// TIA Portal project "PLC_4_LINE4" (V18)

(* hardware
DEVICE "S7-1500/ET200MP station_1"  S7-1500 station
   slot 0: "Rail_0"  Rack  6ES7 590-1***0-0AA0
   slot 1: "PLC_4"  CPU 1511-1 PN  6ES7 511-1AK02-0AB0  V2.9
      slot 3: "CPU display_1"  6ES7591-1AA00-0AA0
      slot 32768: "PROFINET interface_1"  X1
         slot 32769: "Port_1"  X1 P1
         slot 32770: "Port_2"  X1 P2
      slot 34817: "Virtual CP interface port_1"  Virtual CP interface port  Virtual CP interface port
   slot 2: "DI 32x24VDC HF_1"  DI 32x24VDC HF  6ES7 521-1BL00-0AB0  V2.2
   slot 3: "DI 32x24VDC HF_2"  DI 32x24VDC HF  6ES7 521-1BL00-0AB0  V2.2
   slot 4: "DQ 32x24VDC/0.5A HF_1"  DQ 32x24VDC/0.5A HF  6ES7 522-1BL01-0AB0  V1.1
*)

// ===== PLC "PLC_4"  CPU 1511-1 PN =====

VAR_GLOBAL   // PLC tag table "Default tag table"
   "Tag_1" AT %I0.3 : Bool;
   "Tag_2" AT %I0.4 : Bool;
   "Tag_3" AT %I0.5 : Bool;
   "Tag_4" AT %I0.0 : Bool;
   "Tag_5" AT %I0.1 : Bool;
   "Tag_6" AT %I2.1 : Bool;
   "Tag_7" AT %I0.7 : Bool;
   "Tag_8" AT %I1.6 : Bool;
   "Tag_9" AT %I1.0 : Bool;
   "Tag_10" AT %I1.1 : Bool;
   "Tag_11" AT %I1.2 : Bool;
   "Tag_12" AT %I1.3 : Bool;
   "Tag_13" AT %I1.4 : Bool;
   "Tag_14" AT %I1.5 : Bool;
   "Tag_15" AT %Q0.4 : Bool;
   "Tag_16" AT %Q0.5 : Bool;
   "Tag_17" AT %Q0.6 : Bool;
   "Tag_18" AT %Q0.7 : Bool;
   "Tag_19" AT %I4.3 : Bool;
   "Tag_20" AT %I4.4 : Bool;
   "Tag_21" AT %I4.5 : Bool;
   "Tag_22" AT %I4.0 : Bool;
   "Tag_23" AT %I4.1 : Bool;
   "Tag_24" AT %I6.1 : Bool;
   "Tag_25" AT %I4.7 : Bool;
   "Tag_26" AT %I4.6 : Bool;
   "Tag_27" AT %I5.0 : Bool;
   "Tag_28" AT %I5.1 : Bool;
   "Tag_29" AT %I5.2 : Bool;
   "Tag_30" AT %I5.3 : Bool;
   "Tag_31" AT %I5.4 : Bool;
   "Tag_32" AT %I5.5 : Bool;
   "Tag_33" AT %Q2.4 : Bool;
   "Tag_34" AT %Q2.5 : Bool;
   "Tag_35" AT %Q2.6 : Bool;
   "Tag_36" AT %Q2.7 : Bool;
END_VAR

TYPE "typeTask"
   STRUCT
      station : Int;
      dwell_s : Int;
      crane : String[4];
      tank_name : String[10];
      prev : Int;
      next : Int;
      status : Int;
   END_STRUCT;
END_TYPE

TYPE "typeCraneData"
   STRUCT
      task_count : Int;
      tasks : Array[1..20] of "typeTask";
      cmd_send : Bool;
      sts_busy : Bool;
      sts_done : Bool;
      sts_step : Int;
      sts_state : Int;
      ls_at : Array[0..20] of Bool;
      ls_dip : Bool;
      ls_up : Bool;
      ls_mid : Bool;
      btn_start : Bool;
      mv_fwd : Bool;
      mv_rev : Bool;
      mv_up : Bool;
      mv_down : Bool;
      estop : Bool;
      auto : Bool;
      cmd_reset : Bool;
      cmd_stop : Bool;
      pos : Array[0..20] of Int;
   END_STRUCT;
END_TYPE

DATA_BLOCK "Crane6Data"   // DB1
{ S7_Optimized_Access := 'TRUE' }
VERSION : 0.1
BEGIN
   pos[0] := 21;
   pos[1] := 20;
   pos[12] := 14;
   pos[13] := 15;
   pos[14] := 16;
   pos[15] := 17;
   pos[16] := 18;
   pos[17] := 19;
   pos[18] := 20;
END_DATA_BLOCK

DATA_BLOCK "Crane7AData"   // DB2
{ S7_Optimized_Access := 'TRUE' }
VERSION : 0.1
BEGIN
   pos[0] := 2;
   pos[1] := 1;
   pos[2] := 3;
   pos[3] := 4;
   pos[4] := 5;
   pos[5] := 6;
   pos[6] := 7;
   pos[7] := 8;
END_DATA_BLOCK

DATA_BLOCK "Crane6_Seq_DB"   // DB3
{ S7_Optimized_Access := 'TRUE' }
VERSION : 0.1
// stored: InstanceOfName CraneSequencer
"CraneSequencer"
BEGIN
END_DATA_BLOCK

DATA_BLOCK "Crane7A_Seq_DB"   // DB4
{ S7_Optimized_Access := 'TRUE' }
VERSION : 0.1
// stored: InstanceOfName CraneSequencer
"CraneSequencer"
BEGIN
END_DATA_BLOCK

FUNCTION_BLOCK "CraneSequencer"   // FB1, SCL
{ S7_Optimized_Access := 'TRUE' }
VERSION : 0.1
   VAR_IN_OUT
      d : "typeCraneData";
   END_VAR
   VAR
      state : Int;
      idx : Int;
      count : Int;
      cur : Int;
      prevSend : Bool;
      tHold : TON_TIME;
      tDwell : TON_TIME;
   END_VAR
   VAR_TEMP
      target : Int;
      arrived : Bool;
   END_VAR
BEGIN
   // ============================================================================
   //  CraneSequencer  —  GENERIC per-crane batch sequencer  (LIBRARY block)
   // ----------------------------------------------------------------------------
   //  ONE function block reused by EVERY crane on EVERY PLC. Call once per scan
   //  from OB1, passing that crane's data block as the InOut #d. No copy, no
   //  find/replace — the crane it drives is chosen entirely by which DB you pass.
   //
   //  Block type : FUNCTION BLOCK (FB), language SCL.
   //  InOut      : d : "typeCraneData"           // the whole crane interface (a DB of this UDT)
   //  Static     : state:Int, idx:Int, count:Int, cur:Int, prevSend:Bool,
   //               tHold:TON_TIME, tDwell:TON_TIME
   //  Temp       : target:Int, arrived:Bool
   //
   //  OB1 (per crane):  CraneSequencer(d := "Crane6Data")   // its own instance DB
   //                    CraneSequencer(d := "Crane7AData")
   //
   //  Stations: 0=Parking  1=Loading  2..N = tanks (tank number + 1).
   //  States : 0 IDLE · 10 GO_LOAD · 20 LOWER_LOAD · 30 WAIT_BTN · 40 LIFT_LOAD
   //           50 GO_TANK · 60 LOWER_TANK · 70 DWELL · 80 LIFT_TANK · 85 GO_PARK · 90 DONE
   //
   //  DIRECTION IS BY PHYSICAL POSITION, NOT STATION NUMBER.
   //  The plant is NOT laid out in station-number order: Parking sits WEST of Loading, and a
   //  downstream crane's Loading is a transfer tank at the far (West) end. So travel direction
   //  is decided from #d.pos[station] — the physical left→right position of each station
   //  (1 = East-most … larger = further West). TravelTo drives WEST (mv_fwd → R-West) toward a
   //  HIGHER pos, EAST (mv_rev → R-East) toward a LOWER pos. The station's arrival switch is still
   //  #d.ls_at[station]. **Set #d.pos[] per crane** — see the PLC's position-map doc.
   //
   //  COMMANDS (app/Manager writes these):
   //    cmd_send  — arm a batch (rising edge, from IDLE).
   //    cmd_stop  — EMERGENCY HOLD: kills all motion immediately, latches state 100 (STOPPED).
   //                Does NOT clear the recipe. Clear it (and Reset) to move again.
   //    cmd_reset — CLEAN/HOME: lift clear → travel to Parking → wipe the recipe → IDLE.
   //                "As if no recipe was sent, crane back at its home." PLC clears cmd_reset when done.
   //  Extra states: 100 STOPPED · 110 RESET_LIFT · 120 RESET_HOME.
   // ============================================================================

   // ---- command overrides (run BEFORE the state machine, highest priority) ----
   IF #d.cmd_stop THEN                       // immediate emergency hold (latched)
       #d.mv_fwd := FALSE;
       #d.mv_rev := FALSE;
       #d.mv_up := FALSE;
       #d.mv_down := FALSE;
       #d.sts_busy := FALSE;
       #state := 100;
   ELSIF #d.cmd_reset AND #state <> 110 AND #state <> 120 THEN   // start homing/clear (if not already)
       // Wipe the recipe IMMEDIATELY (visible at once), then home the crane.
       #d.task_count := 0;
       #d.sts_step := 0;
       #d.sts_done := FALSE;
       #d.cmd_send := FALSE;
       #idx := 0;
       #count := 0;
       #d.sts_busy := TRUE;
       #state := 110;
   END_IF;

   #d.sts_state := #state;

   CASE #state OF
       0:  // IDLE — parked, hoist up, motors off, waiting for a batch.
           #d.mv_fwd := FALSE;
           #d.mv_rev := FALSE;
           #d.mv_up := FALSE;
           #d.mv_down := FALSE;
           #d.sts_busy := FALSE;
           #d.sts_step := 0;
           IF #d.cmd_send AND NOT #prevSend AND #d.task_count > 0 THEN
               #count := #d.task_count;
               #idx := 1;
               #d.sts_done := FALSE;
               #d.sts_busy := TRUE;
               #state := 10;
           END_IF;

       10: // GO_LOAD — travel to the Loading Area (station 1).
           #d.sts_busy := TRUE;
           #target := 1;
           #arrived := "TravelTo"(target := #d.pos[#target], cur := #d.pos[#cur],
                                  atTarget := #d.ls_at[#target],
                                  fwd => #d.mv_fwd, rev => #d.mv_rev);
           IF #arrived THEN
               #cur := #target;
               #d.mv_fwd := FALSE;
               #d.mv_rev := FALSE;
               #state := 20;
           END_IF;

       20: // LOWER_LOAD — lower the hoist until the dip limit switch is made.
           #d.mv_up := FALSE;
           #d.mv_down := TRUE;
           IF #d.ls_dip THEN
               #d.mv_down := FALSE;
               #state := 30;
           END_IF;

       30: // WAIT_BTN — operator loads material, then HOLDS btn_start for 3 s.
           #tHold(IN := #d.btn_start,
                  PT := T#3S);
           IF #tHold.Q THEN
               #state := 40;
           END_IF;

       40: // LIFT_LOAD — raise the hoist clear before travelling.
           #d.mv_down := FALSE;
           #d.mv_up := TRUE;
           IF #d.ls_up THEN
               #d.mv_up := FALSE;
               #state := 50;
           END_IF;

       50: // GO_TANK — travel to THIS task's tank station (TravelTo reverses if lower).
           #d.sts_step := #idx;
           #d.tasks[#idx].status := 1;                  // running
           #target := #d.tasks[#idx].station;
           #arrived := "TravelTo"(target := #d.pos[#target], cur := #d.pos[#cur],
                                  atTarget := #d.ls_at[#target],
                                  fwd => #d.mv_fwd, rev => #d.mv_rev);
           IF #arrived THEN
               #cur := #target;
               #d.mv_fwd := FALSE;
               #d.mv_rev := FALSE;
               #state := 60;
           END_IF;

       60: // LOWER_TANK — dip into the tank until the dip limit switch is made.
           #d.mv_up := FALSE;
           #d.mv_down := TRUE;
           IF #d.ls_dip THEN
               #d.mv_down := FALSE;
               #state := 70;
           END_IF;

       70: // DWELL — hold in the tank for this task's dwell_s seconds.
           #tDwell(IN := TRUE,
                   PT := DINT_TO_TIME(INT_TO_DINT(#d.tasks[#idx].dwell_s) * 1000));
           IF #tDwell.Q THEN
               #tDwell(IN := FALSE,
                       PT := T#0S);        // reset the timer for the next tank
               #state := 80;
           END_IF;

       80: // LIFT_TANK — lift out, mark the task done, advance or finish.
           #d.mv_down := FALSE;
           #d.mv_up := TRUE;
           IF #d.ls_up THEN
               #d.mv_up := FALSE;
               #d.tasks[#idx].status := 2;              // done
               IF #idx < #count THEN
                   #idx := #idx + 1;
                   #state := 50;                        // next tank
               ELSE
                   #state := 85;                        // all tanks done
               END_IF;
           END_IF;

       85: // GO_PARK — return home to Parking (station 0).
           #target := 0;
           #arrived := "TravelTo"(target := #d.pos[#target], cur := #d.pos[#cur],
                                  atTarget := #d.ls_at[#target],
                                  fwd => #d.mv_fwd, rev => #d.mv_rev);
           IF #arrived THEN
               #cur := #target;
               #d.mv_fwd := FALSE;
               #d.mv_rev := FALSE;
               #state := 90;
           END_IF;

       90: // DONE — raise the done flag, wait for the app to acknowledge (cmd_send → FALSE).
           #d.sts_busy := FALSE;
           #d.sts_done := TRUE;
           IF NOT #d.cmd_send THEN
               #d.sts_done := FALSE;
               #d.sts_step := 0;
               #state := 0;
           END_IF;

       100: // STOPPED — emergency hold. Motors off; leaves only via Reset (cmd_reset).
           #d.mv_fwd := FALSE;
           #d.mv_rev := FALSE;
           #d.mv_up := FALSE;
           #d.mv_down := FALSE;
           #d.sts_busy := FALSE;

       110: // RESET_LIFT — raise the hoist clear before homing.
           #d.mv_down := FALSE;
           #d.mv_up := TRUE;
           IF #d.ls_up THEN
               #d.mv_up := FALSE;
               #state := 120;
           END_IF;

       120: // RESET_HOME — travel to Parking, then wipe the recipe → IDLE.
           #target := 0;
           #arrived := "TravelTo"(target := #d.pos[#target], cur := #d.pos[#cur],
                                  atTarget := #d.ls_at[#target],
                                  fwd => #d.mv_fwd, rev => #d.mv_rev);
           IF #arrived THEN
               #cur := 0;
               #d.mv_fwd := FALSE;
               #d.mv_rev := FALSE;
               #d.task_count := 0;          // "as if no recipe was sent"
               #d.sts_step := 0;
               #d.sts_done := FALSE;
               #d.sts_busy := FALSE;
               #d.cmd_send := FALSE;
               #d.cmd_reset := FALSE;      // handshake: reset complete
               #idx := 0;
               #count := 0;
               #state := 0;                 // IDLE
           END_IF;
   END_CASE;

   #prevSend := #d.cmd_send;   // edge memory (runs every scan, after the CASE)
END_FUNCTION_BLOCK

FUNCTION "IOMap" : Void   // FC1, SCL
{ S7_Optimized_Access := 'TRUE' }
VERSION : 0.1
BEGIN
   // ============================================================================
   //  IOMap  —  PLC_4 (Line 4, cranes 6 & 7A)  —  real %I/%Q  ↔  crane DB mirrors
   // ----------------------------------------------------------------------------
   //  Block type : FUNCTION (FC), language SCL, return type Void, NO parameters.
   //  Call it FIRST in OB1 (before the crane sequencers) so inputs are fresh and
   //  the motor bits the sequencers set this scan reach %Q the same scan.
   //
   //  Addresses are taken verbatim from docs/plc/plant-panel-layout.md (PLC_4).
   //  The %I/%Q addresses must match the hardware I/O module addresses in the PLC
   //  tag table / device config.
   //
   //  Station map: 0=Parking  1=Loading  s = tank.number + 1  (line-wide numbering).
   // ============================================================================

   // ============================ CRANE 6  (Crane6Data) ==========================
   //  Crane 6 is DOWNSTREAM (no loading bay) — it picks material up at TRVL-4A, so
   //  Loading (station 1) is mapped to the same TRVL-4A switch as station 18.
   // --- inputs  %I -> mirror ---
   "Crane6Data".ls_mid := "Tag_1";      // LS_Mid_C6
   "Crane6Data".ls_up := "Tag_2";      // LS_Up_C6
   "Crane6Data".ls_dip := "Tag_3";      // LS_Down_C6
   "Crane6Data".estop := "Tag_4";      // E-Stop_SW_C6   (mirror only; interlock = follow-up)
   "Crane6Data".auto := "Tag_5";      // Auto_SW_C6
   "Crane6Data".btn_start := "Tag_6";      // UP_Pendant_C6  (hold 3 s to start)
   "Crane6Data".ls_at[0] := "Tag_7";      // PRK-4A_C6      (Parking)
   "Crane6Data".ls_at[1] := "Tag_8";      // TRVL-4A_C6     (Loading = transfer pickup)
   "Crane6Data".ls_at[12] := "Tag_9";      // 1-7B_C6   (tank 11 -> station 12)
   "Crane6Data".ls_at[13] := "Tag_10";      // 1-8_C6    (tank 12 -> station 13)
   "Crane6Data".ls_at[14] := "Tag_11";      // 1-9_C6    (tank 13 -> station 14)
   "Crane6Data".ls_at[15] := "Tag_12";      // 1-10A_C6  (tank 14 -> station 15)
   "Crane6Data".ls_at[16] := "Tag_13";      // 1-10B_C6  (tank 15 -> station 16)
   "Crane6Data".ls_at[17] := "Tag_14";      // 1-11_C6   (tank 16 -> station 17)
   "Crane6Data".ls_at[18] := "Tag_8";      // TRVL-4A_C6 (tank 17 -> station 18)
   // --- outputs  mirror -> %Q ---
   "Tag_15" := "Crane6Data".mv_up;          // R-Up-1_C6
   "Tag_16" := "Crane6Data".mv_down;        // R-Down-1_C6
   "Tag_17" := "Crane6Data".mv_rev;         // R-East-1_C6   (East = reverse / left / lower station)
   "Tag_18" := "Crane6Data".mv_fwd;         // R-West-1_C6   (West = forward / right / higher station)

   // ============================ CRANE 7A  (Crane7AData) ========================
   //  Crane 7A is the line ENTRY crane (has LOAD bays). Fully wired from the
   //  Panel_4 drawing: parking + the six entry-tank switches live on input card 2
   //  (%I4.x / %I5.x / %I6.x).
   // --- inputs  %I -> mirror ---
   "Crane7AData".ls_mid := "Tag_19";     // LS_Mid_C7A
   "Crane7AData".ls_up := "Tag_20";     // LS_Up_C7A
   "Crane7AData".ls_dip := "Tag_21";     // LS_Down_C7A
   "Crane7AData".estop := "Tag_22";     // E-Stop_SW_C7A
   "Crane7AData".auto := "Tag_23";     // Auto_SW_C7A
   "Crane7AData".btn_start := "Tag_24";     // UP_Pendant_C7A
   "Crane7AData".ls_at[0] := "Tag_25";     // PRK-4C-C7A   (Parking — crane 7A home)
   "Crane7AData".ls_at[1] := "Tag_26";     // LOAD-4A-C7A  (Loading; LOAD-4B/4C/4D = I6.3/6.4/6.5 extra bays)
   "Crane7AData".ls_at[2] := "Tag_27";     // 1-1A-C7A  (tank 1 -> station 2)
   "Crane7AData".ls_at[3] := "Tag_28";     // 1-1B-C7A  (tank 2 -> station 3)
   "Crane7AData".ls_at[4] := "Tag_29";     // 1-2-C7A   (tank 3 -> station 4)
   "Crane7AData".ls_at[5] := "Tag_30";     // 1-3-C7A   (tank 4 -> station 5)
   "Crane7AData".ls_at[6] := "Tag_31";     // 1-4A-C7A  (tank 5 -> station 6)
   "Crane7AData".ls_at[7] := "Tag_32";     // 1-4B-C7A  (tank 6 -> station 7)
   // --- outputs  mirror -> %Q ---
   "Tag_33" := "Crane7AData".mv_up;         // R-Up-1_C7A
   "Tag_34" := "Crane7AData".mv_down;       // R-Down-1_C7A
   "Tag_35" := "Crane7AData".mv_rev;        // R-East-1_C7A
   "Tag_36" := "Crane7AData".mv_fwd;        // R-West-1_C7A
END_FUNCTION

FUNCTION "TravelTo" : Bool   // FC2, SCL
{ S7_Optimized_Access := 'TRUE' }
VERSION : 0.1
   VAR_INPUT
      target : Int;
      cur : Int;
      atTarget : Bool;
   END_VAR
   VAR_OUTPUT
      fwd : Bool;
      rev : Bool;
   END_VAR
BEGIN
   // TravelTo — pick the travel direction toward a target station.
   // Returns TRUE when the target limit switch is already made (arrived → stop).
   #fwd := FALSE;
   #rev := FALSE;

   IF #atTarget THEN
       ;                       // arrived: leave both motors off
   ELSIF #target > #cur THEN
       #fwd := TRUE;           // higher station number → travel forward
   ELSE
       #rev := TRUE;           // lower station number → travel reverse
   END_IF;

   #TravelTo := #atTarget;
END_FUNCTION

ORGANIZATION_BLOCK "Main"   // OB1, LAD, ProgramCycle
TITLE = "Main Program Sweep (Cycle)"
{ S7_Optimized_Access := 'TRUE' }
VERSION : 0.1
   VAR_INPUT
      Initial_Call : Bool;   // Initial call of this OB
      Remanence : Bool;   // =True, if remanent data are available
   END_VAR
BEGIN

REGION Network 1
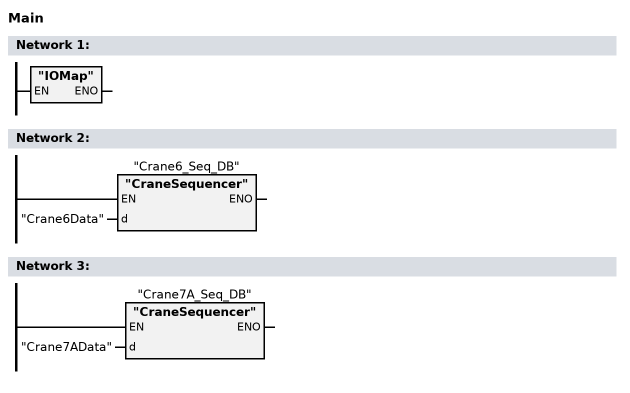
   RUNG wire#powerrail
      "IOMap"()
   END_RUNG
   // the same network as SCL:
   "IOMap"();
END_REGION

REGION Network 2
   RUNG wire#powerrail
      "Crane6_Seq_DB"(d := "Crane6Data")
   END_RUNG
   // the same network as SCL:
   "Crane6_Seq_DB"(d := "Crane6Data");   // "CraneSequencer"
END_REGION

REGION Network 3
   RUNG wire#powerrail
      "Crane7A_Seq_DB"(d := "Crane7AData")
   END_RUNG
   // the same network as SCL:
   "Crane7A_Seq_DB"(d := "Crane7AData");   // "CraneSequencer"
END_REGION
END_ORGANIZATION_BLOCK